(* IEC 61131-3 sources: plc_generation_empirical_study/datasets/packages/internal_v0_1/qualification_only/C10_E01_master_follower_coordination, 1 file *)

(* ---- reference.st ---- *)
FUNCTION_BLOCK C10_E01_master_follower_coordination
VAR_INPUT
    RunRequest : BOOL;
    MasterReady : BOOL;
    FollowerReady : BOOL;
END_VAR
VAR_OUTPUT
    MasterRun : BOOL;
    FollowerRun : BOOL;
END_VAR

MasterRun := RunRequest AND MasterReady;
FollowerRun := RunRequest AND MasterRun AND FollowerReady;

END_FUNCTION_BLOCK
